FUNCTION F_Clamp : LREAL
VAR_INPUT
	fValue	: LREAL;
	fMin	: LREAL;
	fMax	: LREAL;
END_VAR

F_Clamp := MIN(MAX(fValue, fMin), fMax);

END_FUNCTION

(* stored: Version 1.1.0.1
   POU F_Clamp: Id {c2e525fb-4573-4955-b110-db334657dc60}, SpecialFunc None *)
